// Coordinate transforms of an equatorial (HA/Dec) telescope, without axes, clock or comm (IAG50cm#17). The owner sets the
// inputs and calls Target() and Current() in its scan: Target() before it runs its pointing model (which needs
// fHourAngleApparent/fDeclinationApparent), Current() after (it needs the axis positions and the inversion).
// Moved out of IAG50cm's FB_TelescopeControl with the same AstroBROT calls in the same order, and ONE FB_EQ2HOR
// instance for the three conversions to Alt/Az, as there (FB_EQ2HOR keeps state between calls).
// eRefractionMode (IAG50cm#7, #3): OLD gives every AstroBROT call its defaults, as before. NEW passes the weather
// (F_RefractionWeather), takes the slew altitude as observed and publishes the observed sky altitude; the owner then
// runs FB_EqPointing with the same mode and the fRefraction* outputs. fElevationCurrent (the horizon guards) is the
// same in both modes.
FUNCTION_BLOCK FB_RaDecCoordinates
VAR_INPUT
	fJd						: LREAL;		// Julian date, UTC
	fTimeOffset				: LREAL;		// added to fJd for all conversions (TCS time offset)
	fLongitude				: LREAL;		// degrees
	fLatitude				: LREAL;		// degrees
	fAltitude				: LREAL;		// height above sea level, metres
	// target (TCS input)
	fRightAscension			: LREAL;		// ICRS, degrees
	fDeclination			: LREAL;		// ICRS, degrees
	// slew target (TCS input)
	fElevation				: LREAL;		// degrees
	fAzimuth				: LREAL;		// degrees
	// slew target of a SlewHaDec (I_RaDecTelescope.SlewHaDec): while bSlewHaDec, the slew target is this apparent HA/Dec
	// instead of fElevation/fAzimuth, and its ICRS position and Alt/Az are derived from it (IAG50cm X5)
	bSlewHaDec				: BOOL;
	fSlewHaDecHa			: LREAL;		// degrees, apparent
	fSlewHaDecDec			: LREAL;		// degrees, apparent
	// TRUE: the slew altitude is an observed (refracted) one, FALSE: a theoretical one. IAG50cm runs FALSE
	// (IAG50cm#3 decides), AstroBROT's own default and MONET's choice is TRUE.
	bSlewAltIsObserved		: BOOL := TRUE;	// NEW always takes the slew altitude as observed
	eRefractionMode			: E_RefractionMode := E_RefractionMode.OLD;
	stWeather				: ST_Weather;	// live weather (FB_Comm_MQTT_Influx.Weather), used in NEW only
	// axis positions and corrections
	fHourAngleCurrent		: LREAL;		// degrees
	fDeclinationCurrent		: LREAL;		// degrees
	fHourAngleOffset		: LREAL;		// user offset on the sky (cross-declination), degrees
	fDeclinationOffset		: LREAL;		// user offset, degrees
	fHourAngleInversion		: LREAL;		// inverse pointing correction of this scan
	fDeclinationInversion	: LREAL;
	bInversionValid			: BOOL;			// FALSE: the inversion did not converge, keep the last valid correction
END_VAR
VAR_OUTPUT
	// Target()
	fHourAngleApparent		: LREAL;		// apparent hour angle of the target
	fDeclinationApparent	: LREAL;		// apparent declination of the target
	fElevationCalc			: LREAL;		// Alt/Az of the target
	fAzimuthCalc			: LREAL;
	fRightAscensionCalc		: LREAL;		// RA (ICRS) of the slew target
	fDeclinationCalc		: LREAL;		// apparent declination of the slew target, the one the axes are driven to (IAG50cm#239)
	fHourAngleCalc			: LREAL;		// apparent hour angle of the slew target
	fDeclinationCalcIcrs	: LREAL;		// ICRS declination of the slew target (goto coordinates, RaDec)
	fElevationSlew			: LREAL;		// Alt/Az of the slew target: fElevation/fAzimuth, or derived from the SlewHaDec target
	fAzimuthSlew			: LREAL;
	bRefractionNew			: BOOL;			// eRefractionMode = NEW in the last Target()
	bRefractionLiveWeather	: BOOL;			// a live pressure or temperature is used (F_RefractionWeather), NEW only
	fRefractionPressure		: LREAL;		// hPa, 0.0 = estimate; what the AstroBROT calls get (0.0 in OLD)
	fRefractionTemperature	: LREAL;		// deg C
	bRefractionTemperatureSet	: BOOL;
	// Current()
	fRightAscensionCurrentICRS		: LREAL;	// where the axes point, without offsets and pointing correction
	fDeclinationCurrentICRS			: LREAL;
	fRightAscensionCurrentICRScorr	: LREAL;	// where the sky is, with offsets and the inverse pointing correction
	fDeclinationCurrentICRScorr		: LREAL;
	fElevationCurrent		: LREAL;		// Alt/Az of the axes
	fAzimuthCurrent			: LREAL;
	fElevationCurrentSky	: LREAL;		// Alt/Az of the sky position
	fAzimuthCurrentSky		: LREAL;
	fHourAngleInversionHeld		: LREAL;	// the inversion actually used (last valid one)
	fDeclinationInversionHeld	: LREAL;
END_VAR
VAR
	fbRaDec2HaDec	: FB_RADEC2HADEC;
	fbEq2Hor		: FB_EQ2HOR;
	fbHor2Eq		: FB_HOR2EQ;
	fbHaDec2RaDec	: FB_HADEC2RADEC;	// also the SlewHaDec target, one instance as in IAG50cm
	fbRaDec2HaDecSlew	: FB_RADEC2HADEC;	// apparent declination of the Alt/Az slew target (IAG50cm#239)
END_VAR

// the work is in Target() and Current(), the owner decides where in its scan they run

// Apparent HA/Dec of the target, its Alt/Az (to check if it is on the sky or in the ground) and the RA/Dec/HA of the slew target
// (Alt/Az, or the apparent HA/Dec of a SlewHaDec).
METHOD Target
VAR
END_VAR
// the refraction mode of this cycle; the weather only enters in NEW
bRefractionNew := eRefractionMode = E_RefractionMode.NEW;
bRefractionLiveWeather := F_RefractionWeather(
	stWeather		:= stWeather,
	fSiteAltitude	:= fAltitude,
	fPressure		=> fRefractionPressure,
	fTemperature	=> fRefractionTemperature,
	bTemperatureSet	=> bRefractionTemperatureSet);
IF NOT bRefractionNew THEN
	bRefractionLiveWeather := FALSE;
	fRefractionPressure := 0.0;	// the AstroBROT defaults: OLD stays as it was
	fRefractionTemperature := 0.0;
	bRefractionTemperatureSet := FALSE;
END_IF

fbRaDec2HaDec(
	ra := fRightAscension,
	dec := fDeclination,
	lon := fLongitude,
	JD := fJd + fTimeOffset,
	ha_out => fHourAngleApparent,
	dec_out => fDeclinationApparent);
fbEq2Hor(
	ra := fRightAscension,
	dec := fDeclination,
	lon := fLongitude,
	lat := fLatitude,
	altitude := fAltitude,
	JD := fJd + fTimeOffset,
	refract_to_observed := TRUE,
	pressure := fRefractionPressure,
	temperature := fRefractionTemperature,
	temperature_set := bRefractionTemperatureSet,
	alt => fElevationCalc,
	az => fAzimuthCalc);
IF bSlewHaDec THEN
	// SlewHaDec (IAG50cm X5): the target is the apparent HA/Dec itself. Its ICRS position and horizontal coordinates are
	// derived from it, so that the horizon and pole guards, the dome azimuth and the goto coordinates follow the same target.
	fHourAngleCalc := fSlewHaDecHa;
	fDeclinationCalc := fSlewHaDecDec;
	fbHaDec2RaDec(
		ha := fSlewHaDecHa,
		dec := fSlewHaDecDec,
		jd := fJd + fTimeOffset,
		lon := fLongitude,
		ra_out => fRightAscensionCalc,
		dec_out => fDeclinationCalcIcrs);
	fbEq2Hor(
		ra := fRightAscensionCalc,
		dec := fDeclinationCalcIcrs,
		lon := fLongitude,
		lat := fLatitude,
		altitude := fAltitude,
		refract_to_observed := bRefractionNew,	// OLD: FALSE, as in IAG50cm; NEW: the observed altitude, as the published one
		pressure := fRefractionPressure,
		temperature := fRefractionTemperature,
		temperature_set := bRefractionTemperatureSet,
		JD := fJd + fTimeOffset,
		alt => fElevationSlew,
		az => fAzimuthSlew);
ELSE
	fbHor2Eq(
		alt := fElevation,
		az := fAzimuth,
		jd := fJd + fTimeOffset,
		lat := fLatitude,
		lon := fLongitude,
		altitude := fAltitude,
		alt_is_observed := bSlewAltIsObserved OR bRefractionNew,
		pressure := fRefractionPressure,
		temperature := fRefractionTemperature,
		temperature_set := bRefractionTemperatureSet,
		ra => fRightAscensionCalc,
		dec => fDeclinationCalcIcrs,
		ha => fHourAngleCalc);
	// FB_HOR2EQ returns the apparent hour angle but the J2000 declination: the axes are driven in apparent HA/Dec, so take
	// the apparent declination of the same point (IAG50cm#239: mixing the two put the target 0.054 deg off in altitude)
	fbRaDec2HaDecSlew(
		ra := fRightAscensionCalc,
		dec := fDeclinationCalcIcrs,
		lon := fLongitude,
		JD := fJd + fTimeOffset,
		dec_out => fDeclinationCalc);
	fElevationSlew := fElevation;
	fAzimuthSlew := fAzimuth;
END_IF
END_METHOD

// Where the axes point and where that is on the sky: ICRS raw and corrected, Alt/Az raw and sky.
// Needs Target() of the same scan (the HA offset on the axis uses fDeclinationApparent).
METHOD Current
VAR
END_VAR
// near the horizon the inversion is chaotic and does not converge: keep the last trustworthy correction
IF bInversionValid THEN
	fHourAngleInversionHeld := fHourAngleInversion;
	fDeclinationInversionHeld := fDeclinationInversion;
END_IF

// transform from apparent to icrs
fbHaDec2RaDec(
	ha := fHourAngleCurrent,
	dec := fDeclinationCurrent,
	jd := fJd + fTimeOffset,
	lon := fLongitude,
	ra_out => fRightAscensionCurrentICRS,
	dec_out => fDeclinationCurrentICRS);
fbHaDec2RaDec(
	ha := fHourAngleCurrent - fHourAngleInversionHeld - F_HourAngleOffsetOnAxis(fHourAngleOffset, fDeclinationApparent),
	dec := fDeclinationCurrent - fDeclinationInversionHeld - fDeclinationOffset,
	jd := fJd + fTimeOffset,
	lon := fLongitude,
	ra_out => fRightAscensionCurrentICRScorr,
	dec_out => fDeclinationCurrentICRScorr);

// to Alt/Az
fbEq2Hor(
	ra := fRightAscensionCurrentICRS,
	dec := fDeclinationCurrentICRS,
	lon := fLongitude,
	lat := fLatitude,
	altitude := fAltitude,
	refract_to_observed := FALSE,	// both modes: the horizon guards keep their physical position (IAG50cm#7)
	pressure := 0.0,
	temperature := 0.0,
	temperature_set := FALSE,
	JD := fJd + fTimeOffset,
	alt => fElevationCurrent,
	az => fAzimuthCurrent);
fbEq2Hor(
	ra := fRightAscensionCurrentICRScorr,
	dec := fDeclinationCurrentICRScorr,
	lon := fLongitude,
	lat := fLatitude,
	altitude := fAltitude,
	// OLD: FALSE as before. NEW: the corrected position is geometric, the published altitude is the observed one, as the
	// commanded altitude of an Alt/Az slew (IAG50cm#3, #7)
	refract_to_observed := bRefractionNew,
	pressure := fRefractionPressure,
	temperature := fRefractionTemperature,
	temperature_set := bRefractionTemperatureSet,
	JD := fJd + fTimeOffset,
	alt => fElevationCurrentSky,
	az => fAzimuthCurrentSky);
END_METHOD

END_FUNCTION_BLOCK

(* stored: Version 1.1.0.1, ProductVersion 3.1.4024.15
   POU FB_RaDecCoordinates: Id {f96385ec-2b4a-4c27-b494-c794cd2acaf2}, SpecialFunc None
   Method Target: Id {7b36f19e-4b13-4d56-90e2-22d3be9fa356}
   Method Current: Id {a917cf6a-ee29-4454-a35e-971ad1558fbd} *)
